{region 'Documentation'}
(*!
<summary>Request-only I_RunControl double; counts calls without simulating lifecycle behavior.</summary>
*)
{endregion}
FUNCTION_BLOCK RunControlRequestRecorder IMPLEMENTS I_RunControl
VAR
    FStartCount : UINT;
    FAbortCount : UINT;
    FResetCount : UINT;
    FStatus : ST_RunControlStatus;
END_VAR

{region 'Documentation'}
(*!
<summary>Passive AbortCount observation for the command-adapter tests.</summary>
*)
{endregion}
{attribute 'monitoring' := 'call'}
PROPERTY PUBLIC AbortCount : UINT //! Passive AbortCount observation for the command-adapter tests.
GET // PUBLIC
AbortCount := FAbortCount;
END_GET
END_PROPERTY

{region 'Documentation'}
(*!
<summary>Clears recorded calls without performing lifecycle work.</summary>
*)
{endregion}
METHOD PUBLIC Clear
FStartCount := 0;
FAbortCount := 0;
FResetCount := 0;
END_METHOD

{region 'Documentation'}
(*!
<summary>Passive Name observation for the command-adapter tests.</summary>
*)
{endregion}
{attribute 'monitoring' := 'variable'}
PROPERTY PUBLIC Name : STRING(GVL_Constants.NameLength) //! Passive Name observation for the command-adapter tests.
GET // PUBLIC
Name := 'CommandTarget';
END_GET
END_PROPERTY

{region 'Documentation'}
(*!
<summary>Records a Abort request only; no lifecycle or buffer operations.</summary>
*)
{endregion}
METHOD PUBLIC RequestAbort
FAbortCount := FAbortCount + 1;
END_METHOD

{region 'Documentation'}
(*!
<summary>Records a Reset request only; no lifecycle or buffer operations.</summary>
*)
{endregion}
METHOD PUBLIC RequestReset
FResetCount := FResetCount + 1;
END_METHOD

{region 'Documentation'}
(*!
<summary>Records a Start request only; no lifecycle or buffer operations.</summary>
*)
{endregion}
METHOD PUBLIC RequestStart
FStartCount := FStartCount + 1;
END_METHOD

{region 'Documentation'}
(*!
<summary>Passive ResetCount observation for the command-adapter tests.</summary>
*)
{endregion}
{attribute 'monitoring' := 'call'}
PROPERTY PUBLIC ResetCount : UINT //! Passive ResetCount observation for the command-adapter tests.
GET // PUBLIC
ResetCount := FResetCount;
END_GET
END_PROPERTY

{region 'Documentation'}
(*!
<summary>Passive Result observation for the command-adapter tests.</summary>
*)
{endregion}
{attribute 'monitoring' := 'call'}
PROPERTY PUBLIC Result : E_Result //! Passive Result observation for the command-adapter tests.
GET // PUBLIC
Result := E_Result.NotEvaluated;
END_GET
END_PROPERTY

{region 'Documentation'}
(*!
<summary>Passive StartCount observation for the command-adapter tests.</summary>
*)
{endregion}
{attribute 'monitoring' := 'call'}
PROPERTY PUBLIC StartCount : UINT //! Passive StartCount observation for the command-adapter tests.
GET // PUBLIC
StartCount := FStartCount;
END_GET
END_PROPERTY

{region 'Documentation'}
(*!
<summary>Passive Status observation for the command-adapter tests.</summary>
*)
{endregion}
PROPERTY PUBLIC Status : ST_RunControlStatus //! Passive Status observation for the command-adapter tests.
GET // PUBLIC
Status := FStatus;
END_GET
END_PROPERTY

END_FUNCTION_BLOCK

(* stored: Version 1.1.0.1
   POU RunControlRequestRecorder: Id {e1684c99-fe0c-4f93-9d36-f73c2f3e757a}, SpecialFunc None
   Property AbortCount: Id {49490000-0000-4000-8000-000000000006}
   Get Get: Id {49490000-0000-4000-8000-000000000007}
   Method Clear: Id {49490000-0000-4000-8000-000000000001}
   Property Name: Id {49490000-0000-4000-8000-000000000011}
   Get Get: Id {49490000-0000-4000-8000-000000000012}
   Method RequestAbort: Id {49490000-0000-4000-8000-000000000005}
   Method RequestReset: Id {49490000-0000-4000-8000-000000000008}
   Method RequestStart: Id {49490000-0000-4000-8000-000000000002}
   Property ResetCount: Id {49490000-0000-4000-8000-000000000009}
   Get Get: Id {49490000-0000-4000-8000-000000000010}
   Property Result: Id {49490000-0000-4000-8000-000000000013}
   Get Get: Id {49490000-0000-4000-8000-000000000014}
   Property StartCount: Id {49490000-0000-4000-8000-000000000003}
   Get Get: Id {49490000-0000-4000-8000-000000000004}
   Property Status: Id {49490000-0000-4000-8000-000000000015}
   Get Get: Id {49490000-0000-4000-8000-000000000016} *)
